FUNCTION_BLOCK Level_Control_Slider (* Composite Function Block Type *)
  (* Standard: 61499-2 *)
  (* Version 0.0, 12/30/2019, prana, nxtControl GmbH, template *)
  PACKAGE Main;
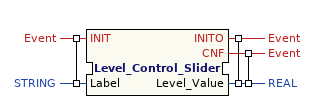
  EVENT_INPUT
    INIT WITH Label; (* Initialization Request *)
  END_EVENT
  EVENT_OUTPUT
    INITO WITH Level_Value; (* Initialization Confirm *)
    CNF WITH Level_Value; (* Execution Confirmation *)
  END_EVENT
  VAR_INPUT
    Label : STRING; (* Input event qualifier *)
  END_VAR
  VAR_OUTPUT
    Level_Value : REAL := 120; (* Output event qualifier *)
  END_VAR
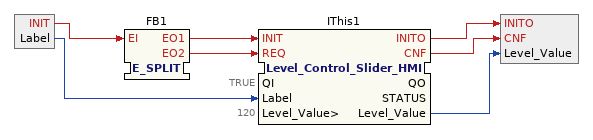
  FBS
    IThis1 : Level_Control_Slider_HMI(Level_Value> := 120, QI := TRUE);
    FB1 : E_SPLIT;
  END_FBS
  EVENT_CONNECTIONS
    INIT TO FB1.EI;
    FB1.EO1 TO IThis1.INIT;
    FB1.EO2 TO IThis1.REQ;
    IThis1.INITO TO INITO;
    IThis1.CNF TO CNF;
  END_CONNECTIONS
  DATA_CONNECTIONS
    Label TO IThis1.Label;
    IThis1.Level_Value TO Level_Value;
  END_CONNECTIONS
END_FUNCTION_BLOCK
